Fanuc KAREL source: KT00506.KL

PROGRAM KT00506
%NOLOCKGROUP
VAR
  P1: XYZWPR
  P2: XYZWPREXT
  OUT: XYZWPREXT
BEGIN
  P1.X = 1.0
    P2.Y = 2.0
  OUT = P1 : P2
END KT00506
